Fanuc KAREL source: kc00029.KL

-- PROVISIONAL review KL for V940-1; original PC SHA256 6736dc628d7e4b2a0b797283939accad2796690bcedb8c95354ad952cfd9ddf9
-- Incomplete behavior may be omitted. Consult companion uncertainty JSON. Do not deploy.
PROGRAM KC00029
%NOLOCKGROUP
BEGIN
  -- V9_ZERO_TABLE_METADATA_HINT layout=0002_ascii; no indexed target words; source/name/runtime held
  -- UNRESOLVED_PC offsets 5-17; opcodes 3F,75
  -- UNRESOLVED_PC offsets 22-106; opcodes 27,22,2A,22,22,22,22,22,22,22,22,22,22,22,22,31
  -- UNRESOLVED_PC offsets 111-115; opcodes 7F
END KC00029
